Fanuc KAREL source: KT00496.KL

PROGRAM KT00496
%NOLOCKGROUP
VAR
  P1: XYZWPR
  P2: POSITION
  OUT: XYZWPREXT
BEGIN
  P1.X = 1.0
  OUT = P1 : P2
END KT00496
